FUNCTION_BLOCK FB_CfcEmpty
VAR_INPUT
END_VAR
VAR_OUTPUT
END_VAR
VAR
END_VAR

END_FUNCTION_BLOCK

(* stored: Version 1.1.0.1, ProductVersion 3.1.4024.12
   POU FB_CfcEmpty: Id {0a1b2c3d-0000-4000-8000-000000000301}, SpecialFunc None *)
